FUNCTION_BLOCK ProcessingComplete (* Composite Function Block Type *)
  (* Standard: 61499-2 *)
  (* Version 0.0, 7/2/2026, template *)
  PACKAGE Main;
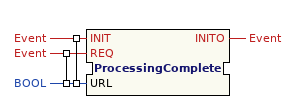
  EVENT_INPUT
    INIT WITH URL; (* Initialization Request *)
    REQ WITH URL; (* Normal Execution Request *)
  END_EVENT
  EVENT_OUTPUT
    INITO; (* Initialization Confirm *)
  END_EVENT
  VAR_INPUT
    URL : BOOL; (* Input event qualifier *)
  END_VAR
END_FUNCTION_BLOCK
